RoboDK station: LineTrack_Station.rdk

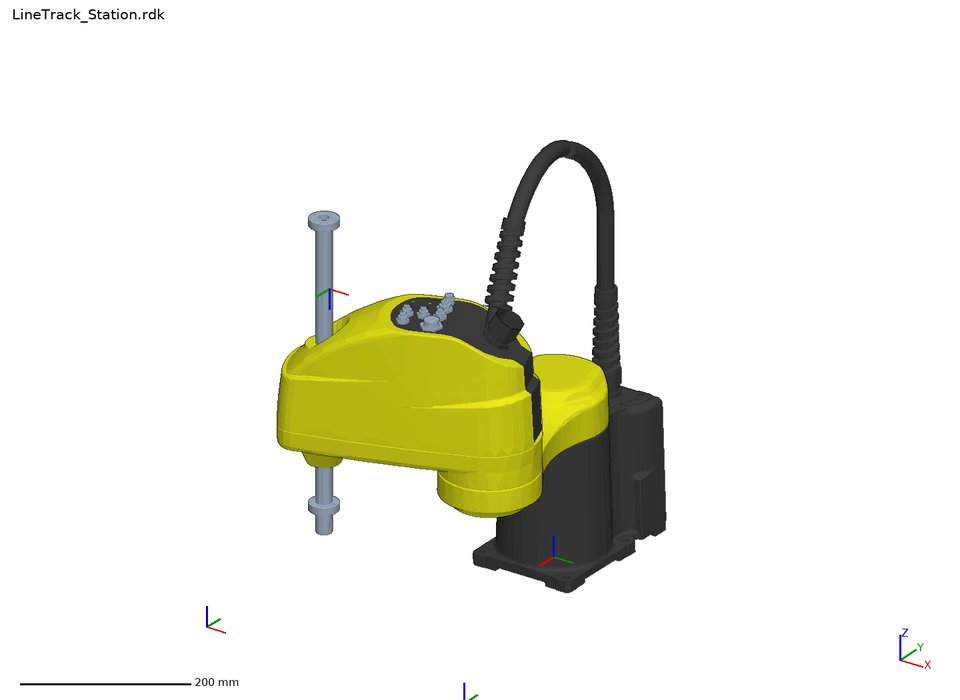
[picture v0: the station drawn from its stored meshes, robots at their saved joint values, targets as dots, program paths as lines]
Station LineTrack_Station (saved by RoboDK 6.0.1). Poses are relative to the parent item; angles as X-Y-Z fixed-axis rotations.
Station parameters (name, value as stored): SICK WL4S Laser Sensor, 0, start_prox, 0
  - frame Fanuc SR-3iA Base at (1214.3, 583.51, 348.22) mm, rotated rx 0 ry 0 rz -90 deg
    - robot Fanuc SR-3iA: 4 axes, payload 3 kg, reach 400 mm, repeatability 0.01 mm, weight 19 kg
        modified DH rows (alpha deg, a mm, theta deg, d mm): 0, 0, 0, 0; 0, 200, 0, 0; 0, 200, 0, 150 linear; 180, 0, 0, 0
        joint limits [-142, -145, -200, -360] to [142, 145, 0, 360]; home [0, 0, 0, 0]; saved at [12.936, -82.426, -50, 69.489]
      - tool Tool 1, TCP at (0, 0, 0) mm
  - frame CamFrame at (1207.08, 136.9, 873.5) mm, rotated rx -180 ry -0.2 rz -0.44 deg
    - camera Camera 1
  - frame Frame 6 at (1375.31, 171.47, 367.78) mm
  - frame Frame 7 at (1050, 111.47, 400) mm
  - frame delete_box_frame at (2400, 111.47, 400) mm
